SUBAPPLICATION FU_Kommando (* Steuerwort vom Web-Dashboard (OPC UA FU1.Kommando) -> 9300H. Genau ein Modbus-Write je Dashboard-Klick, kein zyklisches Nachsenden. *)
  (* Standard: 61499-2; Description: Copyright (c) 2026 Franz Höpfinger This program and the accompanying materials are made available under the terms of the Eclipse Public License 2.0 which is available at https://www.eclipse.org/legal/epl-2.0/ SPDX-License-Identifier: EPL-2.0 *)
  (* Version 1.0, 2026-11-02, Franz Höpfinger, Franz Höpfinger, aus FU_Demo_H300 herausgeloest *)
  PACKAGE FBs::FU_Demo;
  IMPORT FBs::FU_Demo::FU_Demo_Konstanten::FU_MODBUS_KOMMANDO;
  IMPORT FBs::FU_Demo::FU_Demo_Konstanten::FU_KOMMANDO_WEB_READ;
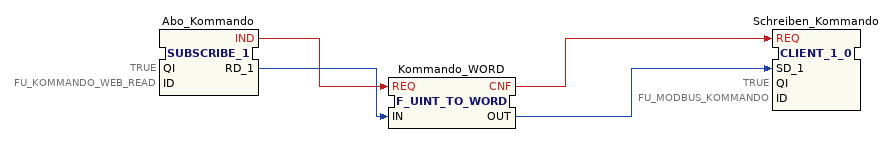
  FBS
    Abo_Kommando : iec61499::net::SUBSCRIBE_1(QI := TRUE, ID := FU_KOMMANDO_WEB_READ);
    Kommando_WORD : iec61131::conversion::F_UINT_TO_WORD; (* typisiert die ANY-Pins: OPC-UA-Knoten wird UInt16, Modbus-Wert WORD *)
    Schreiben_Kommando : iec61499::net::CLIENT_1_0(QI := TRUE, ID := FU_MODBUS_KOMMANDO); (* 9300H Steuerwort *)
  END_FBS
  EVENT_CONNECTIONS
    Abo_Kommando.IND TO Kommando_WORD.REQ;
    Kommando_WORD.CNF TO Schreiben_Kommando.REQ;
  END_CONNECTIONS
  DATA_CONNECTIONS
    Abo_Kommando.RD_1 TO Kommando_WORD.IN;
    Kommando_WORD.OUT TO Schreiben_Kommando.SD_1;
  END_CONNECTIONS
END_SUBAPPLICATION
